Fanuc KAREL source: KA00183.KL

PROGRAM KA00183
%NOLOCKGROUP
VAR
  SRC: ARRAY[4] OF BYTE
  DST: ARRAY[4] OF BOOLEAN
BEGIN
  DST = SRC
END KA00183
